Fanuc KAREL source: KX00032.KL

PROGRAM KX00032
%NOLOCKGROUP
%LOCKGROUP = 1
VAR
  I: INTEGER
  J: INTEGER
  B: BOOLEAN
  F: FILE
  S: STRING[80]
  P: XYZWPR
BEGIN
  I = 1
END KX00032
